(* IEC 61131-3 sources: krc-sample-programs/motor-ramp-alarms-codesys/source/03_States, 2 files *)

(* ---- E_Step.st ---- *)
// The steps. The thousands give the state, the hundreds give the sub-step inside it
// (the four ramp steps and At Speed all belong to Running).
TYPE E_Step :
(
	S0_IDLE      :=    0,	// Idle: powered up and at rest. Goes straight to Not Ready
	S1_NOT_READY := 1000,	// Not Ready: waiting for every permissive, and says which one it is waiting for
	S3_READY     := 3000,	// Ready: waiting for Start
	S4_RAMP_10   := 4000,	// Running: ramping to 10 %
	S4_RAMP_25   := 4100,	// Running: ramping to 25 %
	S4_RAMP_50   := 4200,	// Running: ramping to 50 %
	S4_RAMP_75   := 4300,	// Running: ramping to 75 %
	S4_AT_SPEED  := 4400,	// Running: at speed, 75 %
	S5_STOPPING  := 5000,	// Stopping: speed reference 0, waiting for the motor to stop
	S6_FAULT     := 6000 	// Fault: waiting for the alarm list to clear (Reset clears what it can), then Not Ready
) INT;
END_TYPE

(* ---- CONSTANTS.st ---- *)
// Named numbers the program uses, so no bare number appears in the logic. Constants are all capitals.
VAR_GLOBAL CONSTANT
	SPEED_10           : INT := 10;	// Ramp speed 1, in %
	SPEED_25           : INT := 25;	// Ramp speed 2, in %
	SPEED_50           : INT := 50;	// Ramp speed 3, in %
	SPEED_75           : INT := 75;	// Ramp speed 4 and running speed, in %
	SPEED_STOPPED      : INT := 2;	// At or below this speed, in %, the motor counts as stopped
	SPEED_DEVIATION    : INT := 10;	// At speed, further than this off the reference, in %, is a deviation
	T_SPEED_DEVIATION  : TIME := T#3S;	// ...if it lasts this long
	T_FLASH            : TIME := T#500MS;	// The orange light's flash: this long on, this long off
	AI_FULL_SCALE      : DINT := 32760;	// CC100 analog input at 10 V, in raw counts (WAGO CC100 manual, 9.4)
	AO_FULL_SCALE      : DINT := 32767;	// CC100 analog output count for 10 V (WAGO CC100 manual, 9.4)
	ALARM_COUNT        : INT := 7;	// Lines in the alarm table (GVL_Alarms)
	ALARM_LINES        : INT := 5;	// Alarm lines on the screen
	PERMISSIVE_COUNT   : INT := 4;	// Lines in the permissive table (GVL_Alarms)
	// Where each alarm sits in the alarm table, ALARM level first, so the worst shows at the top
	ALM_ESTOP            : INT := 1;
	ALM_DRIVE_DROPPED    : INT := 2;
	ALM_DRIVE_LOCAL      : INT := 3;
	ALM_RAMP_TIMEOUT     : INT := 4;
	ALM_STOP_TIMEOUT     : INT := 5;
	ALM_SPEED_DEVIATION  : INT := 6;
	ALM_SIM_MODE         : INT := 7;
	// Where each permissive sits in the permissive table, in the order Not Ready names them
	PERM_DRIVE_READY     : INT := 1;
	PERM_DRIVE_REMOTE    : INT := 2;
	PERM_STOP_RELEASED   : INT := 3;
	PERM_MOTOR_STOPPED   : INT := 4;
END_VAR
